FUNCTION_BLOCK TableInit (* Basic Function Block Type *)
  (* Standard: 61499-2 *)
  (* Version 0.0, 7/2/2026, Template *)
  PACKAGE Main;
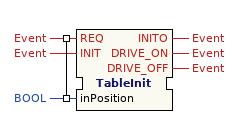
  EVENT_INPUT
    REQ WITH inPosition; (* Normal Execution Request *)
    INIT; (* Initialization Request *)
  END_EVENT
  EVENT_OUTPUT
    INITO; (* Initialization Confirm *)
    DRIVE_ON; (* Execution Confirmation *)
    DRIVE_OFF;
  END_EVENT
  VAR_INPUT
    inPosition : BOOL; (* Input event qualifier *)
  END_VAR
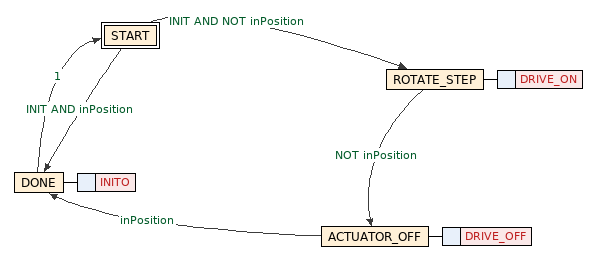
  EC_STATES
    START; (* Initial State *)
    ROTATE_STEP : -> DRIVE_ON;
    ACTUATOR_OFF : -> DRIVE_OFF;
    DONE : -> INITO;
  END_STATES
  EC_TRANSITIONS
    START TO DONE := INIT AND inPosition;
    DONE TO START := 1;
    ROTATE_STEP TO ACTUATOR_OFF := NOT inPosition;
    START TO ROTATE_STEP := INIT AND NOT inPosition;
    ACTUATOR_OFF TO DONE := inPosition;
  END_TRANSITIONS
  ALGORITHM INIT IN ST: (* Initialization algorithm *)
;
  END_ALGORITHM
  ALGORITHM REQ IN ST: (* Normally executed algorithm *)
;
  END_ALGORITHM
END_FUNCTION_BLOCK
